SUBAPPLICATION Uebung_149d (* Übung zu SIZE: zwischen ETP (4000 Byte) und TP (1000 Byte) umschalten *)
  (* Standard: 61499-2; Description: Copyright (c) 2026 Meisterschulen am Ostbahnhof This program and the accompanying materials are made available under the terms of the Eclipse Public License 2.0 which is available at https://www.eclipse.org/legal/epl-2.0/ SPDX-License-Identifier: EPL-2.0 *)
  (* Version 1.0, 2026-11-17, Franz Höpfinger, Meisterschulen am Ostbahnhof, initial API and implementation and/or initial documentation *)
  PACKAGE Uebungen;
  IMPORT Uebungen::const::Uebung_140_149::Etp::LOGIBUS_ADD;
  IMPORT Uebungen::const::Uebung_140_149::Etp::LOGIBUS_FLT;
  IMPORT isobus::pgn::ISOUSERHOME_e::network;
  IMPORT isobus::pgn::ISO_CAN_NODE::NODE1;
  IMPORT isobus::pgn::const::PgnDef::PGN_PDU1_PropA2;
  IMPORT logiBUS::io::DI::logiBUS_DI::Input_I1;
  IMPORT logiBUS::io::DI::logiBUS_DI_Events::BUTTON_SINGLE_CLICK;
  IMPORT logiBUS::io::DI::logiBUS_DI::Input_I2;
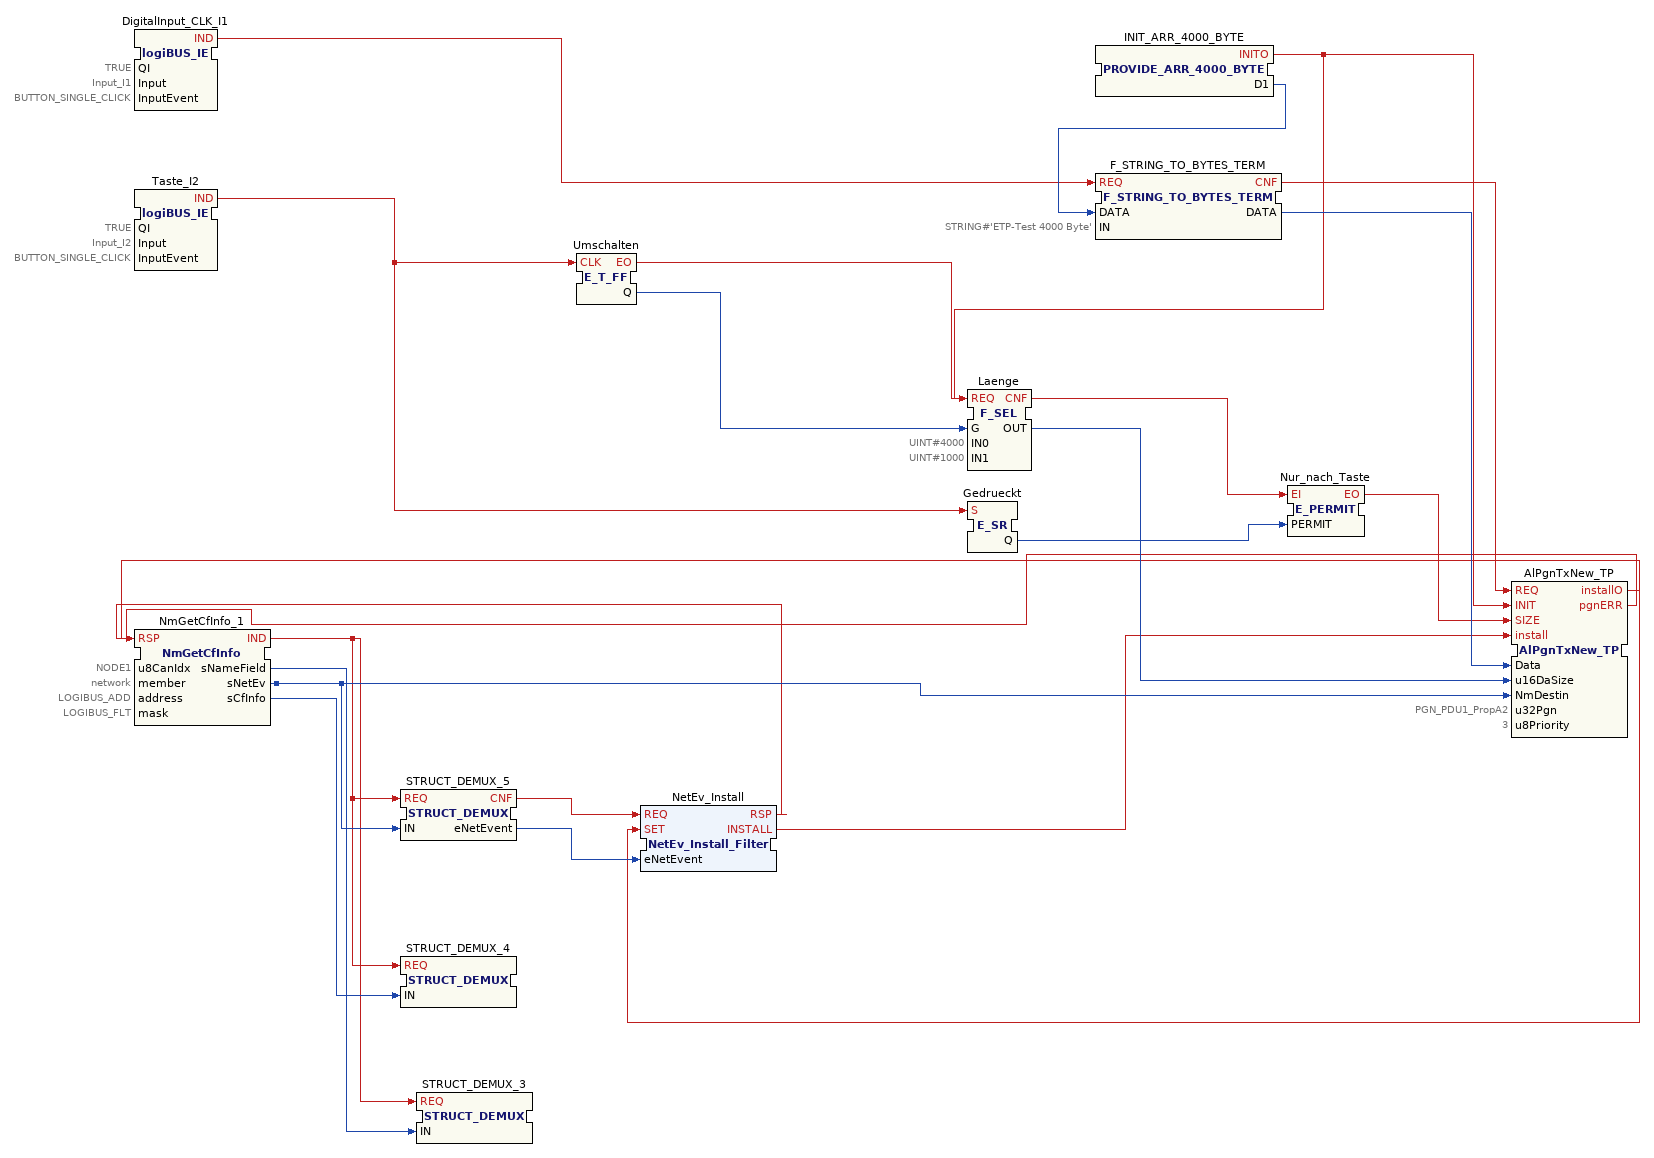
  (* SIZE: zwischen ETP (4000 Byte) und TP (1000 Byte) umschalten, PGN PropA2 0x1EF00 install mit 4000 Byte. I2 Klick schaltet um: 1000 Byte (TP), dann wieder 4000 Byte (ETP). I1 Klick sendet. Der Stack wählt TP oder ETP selbst nach der Länge. Partner wie Übung 149 (Filter LOGIBUS_ADD/LOGIBUS_FLT). Empfänger: Übung 149b, Watch u16DaSize (1000 bzw. 4000). Firmware ab LOGIBUS 24534469 auf BEIDEN Geräten. *)
  FBS
    STRUCT_DEMUX_3 : eclipse4diac::convert::STRUCT_DEMUX; {SET_ATTRIBUTE(StructuredType, isobus::pgn::NAMEFIELD_T)}
    NmGetCfInfo_1 : isobus::pgn::NmGetCfInfo(u8CanIdx := NODE1, member := network, address := LOGIBUS_ADD, mask := LOGIBUS_FLT);
    STRUCT_DEMUX_4 : eclipse4diac::convert::STRUCT_DEMUX; {SET_ATTRIBUTE(StructuredType, isobus::pgn::CF_INFO_T)}
    STRUCT_DEMUX_5 : eclipse4diac::convert::STRUCT_DEMUX; {SET_ATTRIBUTE(StructuredType, isobus::pgn::ISONETEVENT_T)}
    INIT_ARR_4000_BYTE : eclipse4diac::convert::providers::PROVIDE_ARR_4000_BYTE;
    F_STRING_TO_BYTES_TERM : logiBUS::utils::dyn_arr::F_STRING_TO_BYTES_TERM(IN := STRING#'ETP-Test 4000 Byte');
    AlPgnTxNew_TP : isobus::pgn::tx::AlPgnTxNew_TP(u32Pgn := PGN_PDU1_PropA2, u8Priority := 3);
    DigitalInput_CLK_I1 : logiBUS::io::DI::logiBUS_IE(QI := TRUE, Input := Input_I1, InputEvent := BUTTON_SINGLE_CLICK);
    Taste_I2 : logiBUS::io::DI::logiBUS_IE(QI := TRUE, Input := Input_I2, InputEvent := BUTTON_SINGLE_CLICK);
    Umschalten : iec61499::events::E_T_FF;
    Laenge : iec61131::selection::F_SEL(IN0 := UINT#4000, IN1 := UINT#1000); (* Q=FALSE: 4000 Byte ETP (install), Q=TRUE: 1000 Byte TP *)
    Gedrueckt : iec61499::events::E_SR;
    Nur_nach_Taste : iec61499::events::E_PERMIT; (* SIZE erst nach dem ersten Klick *)
  END_FBS
  SUBAPPS
    NetEv_Install : MyLib::sys::NetEv_Install_Filter;
  END_SUBAPPS
  EVENT_CONNECTIONS
    NmGetCfInfo_1.IND TO STRUCT_DEMUX_3.REQ;
    NmGetCfInfo_1.IND TO STRUCT_DEMUX_4.REQ;
    NmGetCfInfo_1.IND TO STRUCT_DEMUX_5.REQ;
    DigitalInput_CLK_I1.IND TO F_STRING_TO_BYTES_TERM.REQ;
    F_STRING_TO_BYTES_TERM.CNF TO AlPgnTxNew_TP.REQ;
    AlPgnTxNew_TP.installO TO NmGetCfInfo_1.RSP;
    AlPgnTxNew_TP.pgnERR TO NmGetCfInfo_1.RSP;
    STRUCT_DEMUX_5.CNF TO NetEv_Install.REQ;
    NetEv_Install.RSP TO NmGetCfInfo_1.RSP;
    AlPgnTxNew_TP.installO TO NetEv_Install.SET;
    INIT_ARR_4000_BYTE.INITO TO Laenge.REQ;
    INIT_ARR_4000_BYTE.INITO TO AlPgnTxNew_TP.INIT;
    Taste_I2.IND TO Gedrueckt.S;
    Taste_I2.IND TO Umschalten.CLK;
    Umschalten.EO TO Laenge.REQ;
    Laenge.CNF TO Nur_nach_Taste.EI;
    Nur_nach_Taste.EO TO AlPgnTxNew_TP.SIZE;
    NetEv_Install.INSTALL TO AlPgnTxNew_TP.install;
  END_CONNECTIONS
  DATA_CONNECTIONS
    NmGetCfInfo_1.sNameField TO STRUCT_DEMUX_3.IN;
    NmGetCfInfo_1.sNetEv TO STRUCT_DEMUX_5.IN;
    NmGetCfInfo_1.sCfInfo TO STRUCT_DEMUX_4.IN;
    INIT_ARR_4000_BYTE.D1 TO F_STRING_TO_BYTES_TERM.DATA;
    F_STRING_TO_BYTES_TERM.DATA TO AlPgnTxNew_TP.Data;
    STRUCT_DEMUX_5.eNetEvent TO NetEv_Install.eNetEvent;
    Gedrueckt.Q TO Nur_nach_Taste.PERMIT;
    Umschalten.Q TO Laenge.G;
    Laenge.OUT TO AlPgnTxNew_TP.u16DaSize;
    NmGetCfInfo_1.sNetEv TO AlPgnTxNew_TP.NmDestin;
  END_CONNECTIONS
END_SUBAPPLICATION
